Staubli VAL3: MoveCirc.pgx

program MoveCirc(num x_nX, num x_nY, num x_nZ, num x_nRx, num x_nRy, num x_nRz, num x_nX2, num x_nY2, num x_nZ2, num x_nRx2, num x_nRy2, num x_nRz2)
begin
  pPointRs.trsf.x = x_nX
  pPointRs.trsf.y = x_nY
  pPointRs.trsf.z = x_nZ
  pPointRs.trsf.rx = x_nRx
  pPointRs.trsf.ry = x_nRy
  pPointRs.trsf.rz = x_nRz
  pPointRs2.trsf.x = x_nX2
  pPointRs2.trsf.y = x_nY2
  pPointRs2.trsf.z = x_nZ2
  pPointRs2.trsf.rx = x_nRx2
  pPointRs2.trsf.ry = x_nRy2
  pPointRs2.trsf.rz = x_nRz2
  movec(pPointRs,pPointRs2,tCurrentTool,mCurrentSpeed)
end
